TYPE ST_NestTracking :
STRUCT
	bPartLoaded       : BOOL;
    bPreviousSensor   : BOOL;
    bPartRemovedPulse : BOOL;
    bPartLoadedPulse  : BOOL;
END_STRUCT
END_TYPE

(* stored: Version 1.1.0.1
   DUT ST_NestTracking: Id {767fb3e8-45a4-4522-8233-925dbd3322a9} *)
